Fanuc KAREL source: kd00064.KL

-- PROVISIONAL review KL for V1013-1; original PC SHA256 5ecba80888d37cb2d3e75f19c963ec0ffbcb76dd3929293276a80650f85bcd22
-- Incomplete behavior may be omitted. Consult companion uncertainty JSON. Do not deploy.
PROGRAM KD00064
%NOLOCKGROUP
VAR
  I : INTEGER
  J : INTEGER
  B : BOOLEAN
  R : REAL
  S : STRING[80]
BEGIN
  -- UNRESOLVED_PC offsets 5-18; opcodes 9D,81,18,9D,1B,9D,12,9C,13,04
  -- UNRESOLVED_PC offsets 23-27; opcodes 7F
END KD00064
